TYPE "LIOLink_3UG4825_typeParam"
TITLE = LIOLink_3UG4825_typeParam
VERSION : 0.1
// Data set (index) 131 (parameters)
   STRUCT
      reserved : Array[0..15] of Byte;   // Reserved
      groupDiagnostics : Bool := TRUE;   // Group diagnostics: Default: true, false; disabled, true: enabled
      groupErrorDiagnostics : Bool := TRUE;   // Group error diagnostics: Default: true, false; disabled, true: enabled
      reserved1 : Bool;   // Reserved
      reserved2 : Bool;   // Reserved
      localLimitChange : Bool := TRUE;   // Local threshold change: Default: true, false; disabled, true: enabled
      localParameterChange : Bool := TRUE;   // Local parameter change: Default: true, false; disabled, true: enabled
      localReset : Bool := TRUE;   // Local reset: Default: true, false; disabled, true: enabled
      retentiveErrorMemory : Bool;   // Retentive error memory: Default: false, false; disabled, true: enabled
      analogValueCoding : Byte := 16#0E;   // Analog value coding: Default: 14, Min: 0(disabled), Max: 255
      reserved3 : Array[18..23] of Byte;   // Reserved
      resetResponse : Byte := 16#01;   // Reset response: Default: 16#01, 16#00: manual, 16#01: automatic
      delayOn : Bool := TRUE;   // ON-delay time (at Power ON): Default: true, false: disabled, true: enabled
      delayOn0 : Bool;   // False
      delayReset : Bool := TRUE;   // ON-delay time (at manual reset): Default: true, false: disabled, true: enabled
      delayReset0 : Bool;   // False
      delayRestart : Bool;   // ON-delay time (at restart): Default: true, false: disabled, true: enabled
      delayRestart0 : Bool;   // False
      reserved4 : Bool;   // Reserved
      reserved5 : Bool;   // Reserved
      delayTime : Int;   // ON-delay time: Resolution: 0.1=1s, Default: 0s, Min: 0.1s or 0s (disabled), Max: 999.9s
      delayTimeTripUp : Int;   // Tripping delay time (in the case of current overshoot): Resolution: 0.1s=1, Default: 0, Min: 0.1s or 0s, Max: 999.9s
      reserved6 : Word;   // Reserved
      tresholdUp : Int := 100;   // Threshold for overshoot: Resolution: 0.01A=1, Default: 1A, Min: 0.03A, Max: 40A
      reserved9 : Word;   // Reserved
      warningTresholdUp : Int := 50;   // Warning threshold for overshoot: Resolution: 0.01A=1, Default: 0,5A, Min: 0.03A or 0A (disabled), Max: 40A
      reserved7 : Array[38..43] of Byte;   // Reserved
      hysteresis : Int := 5;   // Hysteresis: Resolution: Resolution: 1%=1, Default: 5%, Min: 5% or 0% (disabled), Max: 50%
      reserved10 : Byte;   // Reserved
      responseRelay : Byte;   // Relay switching response: Default: 16#00, 16#00: Closed-circuit principle NC, 16#01: Open-circuit principle NO
   END_STRUCT;
END_TYPE

TYPE "LIOLink_3UG4825_typeAll"
TITLE = LIOLink_3UG4825_typeAll
VERSION : 0.1
// Contains all the information about 3UG4825
   STRUCT
      parameterPage0 : "LIOLink_typeParameterPage0";   // ID0: Parameter page 0
      systemCommands : Byte;   // ID2: System Commands (0x80 for device reset, 0x82 for factory reset)
      vendorName : String[11];   // ID16: Vendor name
      vendorText : String[64];   // ID17: Vendor text
      productName : String[64];   // ID18: Product name
      productID : String[14];   // ID19: Product ID
      serialNumber : String[16];   // ID21: Serial number
      hwRevision : String[7];   // ID22: Hardware revision
      fwRevision : String[7];   // ID23: Firmware revision
      appSpecificName : String[32];   // ID24: Application specific name
      diagnostics : "LIOLink_3UG4825_typeDiag";   // ID92: Diagnostics
      measuredValues : "LIOLink_3UG4825_typeMeasure";   // ID94: Measurement values
      parameters : "LIOLink_3UG4825_typeParam";   // ID131: Parameters
   END_STRUCT;
END_TYPE

TYPE "LIOLink_3UG4825_typeDiag"
TITLE = LIOLink_3UG4825_typeDiag
VERSION : 0.1
// Data set (index) 92 - diagnostics
   STRUCT
      reserved : Array[0..15] of Byte;   // Reserved
      ready : Bool;   // Ready
      groupError : Bool;   // Group error
      groupWarning : Bool;   // Group warning
      reserved1 : Bool;   // Reserved
      reserved2 : Bool;   // Reserved
      parameterAssign : Bool;   // Parameter assignment active
      parameterInvalid : Bool;   // Invalid parameter
      internalError : Bool;   // Self-test error/internal error
      reserved3 : Byte;   // Reserved
      errorNumber : Word;   // Parameter error number
      reserved4 : Array[20..25] of Byte;   // Reserved
      delayTimeRunning : Bool;   // ON-delay time running
      delayLevelUp : Bool;   // Tripping delay time running (threshold for overshoot)
      reserved5 : Bool;   // Reserved
      initTimeRunning : Bool;   // Initialization time running after applying the control supply voltage
      reserved6 : Bool;   // Reserved
      reserved7 : Bool;   // Reserved
      reserved8 : Bool;   // Reserved
      reserved9 : Bool;   // Reserved
      levelUp : Bool;   // Threshold for overshoot exceeded
      reserved10 : Bool;   // Reserved
      warningLevelUp : Bool;   // Warning threshold for overshoot exceeded
      reserved11 : Bool;   // Reserved
      reserved12 : Bool;   // Reserved
      reserved13 : Bool;   // Reserved
      reserved14 : Bool;   // Reserved
      reserved15 : Bool;   // Reserved
      wireBreak : Bool;   // Wire break
      shortCircuit : Bool;   // Short-circuit
      rangeOvershoot : Bool;   // Measuring range overshoot
      reserved16 : Bool;   // Reserved
      reserved17 : Bool;   // Reserved
      reserved18 : Bool;   // Reserved
      reserved19 : Bool;   // Reserved
      reserved20 : Bool;   // Reserved
      reserved21 : Byte;   // Reserved
   END_STRUCT;
END_TYPE

// folder: LIOLink/Common/Device-specific data types/SIRIUS/SIRIUS 3UG48/3UG4832

TYPE "LIOLink_3UG4832_typeMeasure"
TITLE = LIOLink_3UG4832_typeMeasure
VERSION : 0.1
// Contains measured value dataset of 3UG4832
   STRUCT
      reserved : Array[0..15] of Byte;   // Reserved
      voltageU1 : Word;   // Voltage
      reserved1 : Array[18..27] of Byte;   // Reserved
   END_STRUCT;
END_TYPE

TYPE "LIOLink_3UG4832_typeParam"
TITLE = LIOLink_3UG4832_typeParam
VERSION : 0.1
// LIOLink_3UG4851_typeParam
   STRUCT
      reserved : Array[0..15] of Byte;   // Reserved
      groupDiagnostics : Bool := TRUE;   // Group diagnostics: Default: true, false; disabled, true: enabled
      groupErrorDiagnostics : Bool := TRUE;   // Group error diagnostics: Default: true, false; disabled, true: enabled
      reserved1 : Bool;   // Reserved
      reserved2 : Bool;   // Reserved
      localLimitChange : Bool := TRUE;   // Local threshold change: Default: true, false; disabled, true: enabled
      localParameterChange : Bool := TRUE;   // Local parameter change: Default: true, false; disabled, true: enabled
      localReset : Bool := TRUE;   // Local reset: Default: true, false; disabled, true: enabled
      retentiveErrorMemory : Bool;   // Retentive error memory: Default: false, false; disabled, true: enabled
      analogValueCoding : Byte := 16#2C;   // Analog value coding: Default: 44, Min: 0(disabled), Max: 255
      reserved3 : Array[18..23] of Byte;   // Reserved
      resetResponse : Byte := 16#01;   // Reset response: Default: 16#01, 16#00: manual, 16#01: automatic
      delayOn : Bool := TRUE;   // ON-delay time (at Power ON): Default: true, false: disabled, true: enabled
      delayOn0 : Bool;   // False
      delayReset : Bool := TRUE;   // ON-delay time (at manual reset): Default: true, false: disabled, true: enabled
      delayReset0 : Bool;   // False
      reserved6 : Bool;   // Reserved
      reserved9 : Bool;   // Reserved
      reserved4 : Bool;   // Reserved
      reserved5 : Bool;   // Reserved
      delayTime : Int := 0;   // ON-delay time: Resolution: 0.1=1s, Default: 0s, Min: 0.1s or 0s (disabled), Max: 999.9s
      delayTimeTripUp : Int;   // Tripping delay time (in the case of voltage overshoot): Resolution: 0.1s=1, Default: 0, Min: 0.1s or 0s, Max: 999.9s
      delayTimeTripDown : Int;   // Tripping delay time (in the case of voltage undershoot): Resolution: 0.1s=1, Default: 0, Min: 0.1s or 0s, Max: 999.9s
      tresholdUp : Int := 3000;   // Threshold for overshoot: Resolution: 0.1V=1, Default: 300, Min: 10V or 0V (disabled), Max: 600V
      tresholdDown : Int := 2000;   // Threshold for undershoot: Resolution: 0.1V=1, Default: 200, Min: 10V or 0V (disabled), Max: 600V
      warningTresholdUp : Int := 3000;   // Warning threshold for overshoot: Resolution: 0.1V=1, Default: 300, Min: 10V or 0V (disabled), Max: 600V
      warningTresholdDown : Int := 2000;   // Warning threshold for undershoot: Resolution: 0.1V=1, Default: 200, Min: 10V or 0V (disabled), Max: 600V
      reserved7 : Array[40..43] of Byte;   // Reserved
      hysteresis : Int := 50;   // Hysteresis: Resolution: 0.1V=1, Default: 5V, Min: 0.1V or 0V (disabled), Max: 300V
      responseRelay : Byte;   // Relay switching response: Default: 16#00, 16#00: Closed-circuit principle NC, 16#01: Open-circuit principle NO
      reserved8 : Byte;   // Reserved
   END_STRUCT;
END_TYPE

TYPE "LIOLink_3UG4832_typeDiag"
TITLE = LIOLink_3UG4832_typeDiag
VERSION : 0.1
// Data set (index) 92 - diagnostics
   STRUCT
      reserved : Array[0..15] of Byte;   // Reserved
      ready : Bool;   // Read
      groupError : Bool;   // Group error
      groupWarning : Bool;   // Group warning
      reserved1 : Bool;   // Reserved
      reserved2 : Bool;   // Reserved
      parameterAssign : Bool;   // Parameter assignment active
      parameterInvalid : Bool;   // Invalid parameter
      internalError : Bool;   // Self-test error/internal error
      reserved3 : Byte;   // Reserved
      errorNumber : Word;   // Parameter error number
      reserved4 : Array[20..25] of Byte;   // Reserved
      delayTimeRunning : Bool;   // ON-delay time running
      delayLevelUp : Bool;   // Tripping delay time running (threshold for overshoot)
      delayLevelDown : Bool;   // Tripping delay time running (threshold for undershoot)
      reserved5 : Bool;   // Reserved
      reserved6 : Bool;   // Reserved
      reserved7 : Bool;   // Reserved
      reserved8 : Bool;   // Reserved
      reserved9 : Bool;   // Reserved
      levelUp : Bool;   // Threshold for overshoot exceeded
      levelDown : Bool;   // Threshold for undershoot violated
      warningLevelUp : Bool;   // Warning threshold for overshoot exceeded
      warningLevelDown : Bool;   // Warning threshold for undershoot violated
      reserved10 : Bool;   // Reserved
      reserved11 : Bool;   // Reserved
      reserved12 : Bool;   // Reserved
      reserved13 : Bool;   // Reserved
   END_STRUCT;
END_TYPE

TYPE "LIOLink_3UG4832_typeAll"
TITLE = LIOLink_3UG4832_typeAll
VERSION : 0.1
// Contains all the information about 3UG4832
   STRUCT
      parameterPage0 : "LIOLink_typeParameterPage0";   // ID0: Parameter page 0
      systemCommands : Byte;   // ID2: System Commands (0x80 for device reset, 0x82 for factory reset)
      vendorName : String[11];   // ID16: Vendor name
      vendorText : String[64];   // ID17: Vendor text
      productName : String[64];   // ID18: Product name
      productID : String[14];   // ID19: Product ID
      hwRevision : String[7];   // ID22: Hardware revision
      fwRevision : String[7];   // ID23: Firmware revision
      appSpecificName : String[32];   // ID24: Application specific name
      diagnostics : "LIOLink_3UG4832_typeDiag";   // ID92: Diagnostics
      measuredValues : "LIOLink_3UG4832_typeMeasure";   // ID94: Measurement values
      parameters : "LIOLink_3UG4832_typeParam";   // ID131: Parameters
   END_STRUCT;
END_TYPE

// folder: LIOLink/Common/Device-specific data types/SIRIUS/SIRIUS 3UG48/3UG4841

TYPE "LIOLink_3UG4841_typeMeasure"
TITLE = LIOLink_3UG4841_typeMeasure
VERSION : 0.1
// Data set (index) 94 (measured values)
   STRUCT
      reserved : Array[0..15] of Byte;   // Reserved
      valueCosPhiPa : Word;   // Cos Phi Value (PA) Min:0 Max:0,99
      currentActivePa : Word;   // Active current Ir/Ires (PA) Min:0,2A Max:10A
      currentApparentPa : Word;   // Apparent current Is (PA) Min:0,2A Max:10A
      voltageActivePa : Word;   // Active voltage U (PA) Min:30V Max:690V
      powerActivePa : Word;   // Active power Pw (PA) Min:6W Max:6900W
      reserved1 : Array[26..29] of Byte;   // Reserved
      currentActive : DWord;   // Active current Ir/Ires (PA) Min:0,2A Max:10A
      currentApparent : DWord;   // Apparent current Is Min:0,2A Max:10A
      powerActive : DWord;   // Active power Pw Min:6W Max:6900W
      reserved2 : Array[42..49] of Byte;   // Reserved
   END_STRUCT;
END_TYPE

TYPE "LIOLink_3UG4841_typeParam"
TITLE = LIOLink_3UG4841_typeParam
VERSION : 0.1
// Data set (index) 131 (parameters)
   STRUCT
      reserved : Array[0..15] of Byte;   // Reserved
      groupDiagnostics : Bool := TRUE;   // Group diagnostics: Default: true, false; disabled, true: enabled
      groupErrorDiagnostics : Bool := TRUE;   // Group error diagnostics: Default: true, false; disabled, true: enabled
      reserved1 : Bool;   // Reserved
      reserved2 : Bool;   // Reserved
      localLimitChange : Bool := TRUE;   // Local threshold change: Default: true, false; disabled, true: enabled
      localParameterChange : Bool := TRUE;   // Local parameter change: Default: true, false; disabled, true: enabled
      localReset : Bool := TRUE;   // Local reset: Default: true, false; disabled, true: enabled
      retentiveErrorMemory : Bool;   // Retentive error memory: Default: false, false; disabled, true: enabled
      analogValueCoding : Byte := 16#2B;   // Analog value coding: Default: 43, Min: 0(disabled), Max: 255
      reserved3 : Array[18..23] of Byte;   // Reserved
      resetResponse : Byte := 16#01;   // Reset response: Default: 16#01, 16#00: manual, 16#01: automatic
      delayOn : Bool := TRUE;   // ON-delay time (at Power ON): Default: true, false: disabled, true: enabled
      delayOn0 : Bool;   // False
      delayReset : Bool := TRUE;   // ON-delay time (at manual reset): Default: true, false: disabled, true: enabled
      delayReset0 : Bool;   // False
      delayRestart : Bool;   // ON-delay time (at restart): Default: true, false: disabled, true: enabled
      delayRestart0 : Bool;   // False
      reserved4 : Bool;   // Reserved
      reserved5 : Bool;   // Reserved
      delayTime : Int;   // ON-delay time: Resolution: 0.1=1s, Default: 0s, Min: 0.1s or 0s (disabled), Max: 999.9s
      delayTimeCosPhiTripUp : Int;   // Tripping delay time (in the case of overshoot of the cos phi value): Resolution: 0.1s=1, Default: 0, Min: 0.1s or 0s, Max: 999.9s
      delayTimeCosPhiTripDown : Int;   // Tripping delay time (in the case of undershoot of the cos phi value): Resolution: 0.1s=1, Default: 0, Min: 0.1s or 0s, Max: 999.9s
      delayTimeCurrentTripUp : Int;   // Tripping delay time (in the case of active current overshoot): Resolution: 0.1s=1, Default: 0, Min: 0.1s or 0s, Max: 999.9s
      delayTimeCurrentTripDown : Int;   // Tripping delay time (in the case of active current undershoot): Resolution: 0.1s=1, Default: 0, Min: 0.1s or 0s, Max: 999.9s
      tresholdCosPhiUp : Byte := 16#32;   // Threshold for overshoot of the cos phi value: Resolution: 0.01=1, Default: 0.5, Min: 0.01 or 0 (disabled), Max: 0.99
      tresholdCosPhiDown : Byte := 16#14;   // Threshold for undershoot of the cos phi value: Resolution: 0.01=1, Default: 0.2, Min: 0.01 or 0 (disabled), Max: 0.99
      tresholdCurrentUp : DInt := 30;   // Threshold for overshoot of the active current value: Resolution: 0.1A=1, Default: 3A, Min: 0.2A or 0A (disabled), Max: 10A
      tresholdCurrentDown : DInt := 10;   // Threshold for undershoot of the active current value: Resolution: 0.1A=1, Default: 1A, Min: 0.2A or 0A (disabled), Max: 10A
      warningTresholdCosPhiUp : Byte := 16#32;   // Warning threshold for overshoot: Resolution: 0.01A=1, Default: 2.5A, Min: 0.05A or 0A (disabled), Max: 10A
      warningTresholdCosPhiDown : Byte := 16#14;   // Warning threshold for undershoot: Resolution: 0.01A=1, Default: 1.5A, Min: 0.05A or 0A (disabled), Max: 10A
      warningTresholdCurrentUp : DInt := 30;   // Warning threshold for overshoot of the active current value: Resolution: 0.1A=1, Default: 3A, Min: 0.2A or 0A (disabled), Max: 10A
      warningTresholdCurrentDown : DInt := 10;   // Warning threshold for undershoot of the active current value: Resolution: 0.1A=1, Default: 1A, Min: 0.2A or 0A (disabled), Max: 10A
      reserved6 : Array[56..65] of Byte;   // Reserved
      hysteresisCosPhi : Byte := 16#0A;   // Hysteresis (cos phi): Resolution: 0.01=1, Default: 0.1, Min: 0.1 or 0 (disabled), Max: 0.2
      reserved7 : Byte;   // Reserved
      hysteresisCurrent : DInt := 5;   // Hysteresis (active current): Resolution: 0.1A=1, Default: 0,5A, Min: 0.1A or 0A (disabled), Max: 3A
      responseRelay : Byte;   // Relay switching response: Default: 16#00, 16#00: Closed-circuit principle NC, 16#01: Open-circuit principle NO
      reserved8 : Byte;   // Reserved
   END_STRUCT;
END_TYPE

TYPE "LIOLink_3UG4841_typeDiag"
TITLE = LIOLink_3UG4841_typeDiag
VERSION : 0.1
// Data set (index) 92 - diagnostics
   STRUCT
      reserved : Array[0..15] of Byte;   // Reserved
      ready : Bool;   // Ready
      groupError : Bool;   // Group error
      groupWarning : Bool;   // Group warning
      reserved1 : Bool;   // Reserved
      reserved2 : Bool;   // Reserved
      parameterAssign : Bool;   // Parameter assignment active
      parameterInvalid : Bool;   // Invalid parameter
      internalError : Bool;   // Self-test error/internal error
      reserved3 : Byte;   // Reserved
      errorNumber : Word;   // Parameter error number
      reserved4 : Array[20..25] of Byte;   // Reserved
      delayTimeRunning : Bool;   // ON-delay time running
      delayCosPhiUp : Bool;   // Tripping delay time running (threshold for overshoot: cos phi value)
      delayLCosPhiDown : Bool;   // Tripping delay time running (threshold for undershoot: cos phi value)
      delayCurrentUp : Bool;   // Tripping delay time running (threshold for overshoot: active current value)
      delayCurrentDown : Bool;   // Tripping delay time running (threshold for undershoot: active current value)
      reserved5 : Bool;   // Reserved
      reserved6 : Bool;   // Reserved
      reserved7 : Bool;   // Reserved
      cosPhiUp : Bool;   // Threshold value for overshoot exceeded (cos phi value)
      cosPhiDown : Bool;   // Threshold value for undershoot violated (cos phi value)
      currentUp : Bool;   // Threshold for overshoot exceeded (active current value)
      currentDown : Bool;   // Threshold for undershoot violated (active current value)
      warningCosPhiUp : Bool;   // Warning threshold for overshoot exceeded (cos phi value)
      warningCosPhiDown : Bool;   // Warning threshold for undershoot violated (cos phi value)
      warningCurrentUp : Bool;   // Warning threshold for overshoot exceeded (active current value)
      warningCurrentDown : Bool;   // Warning threshold for undershoot violated (active current value)
      reserved8 : Word;   // Reserved
   END_STRUCT;
END_TYPE

TYPE "LIOLink_3UG4841_typeAll"
TITLE = LIOLink_3UG4841_typeAll
VERSION : 0.1
// Contains all the information about 3UG4841
   STRUCT
      parameterPage0 : "LIOLink_typeParameterPage0";   // ID0: Parameter page 0
      systemCommands : Byte;   // ID2: System Commands (0x80 for device reset, 0x82 for factory reset)
      vendorName : String[11];   // ID16: Vendor name
      vendorText : String[64];   // ID17: Vendor text
      productName : String[64];   // ID18: Product name
      productID : String[14];   // ID19: Product ID
      hwRevision : String[7];   // ID22: Hardware revision
      fwRevision : String[7];   // ID23: Firmware revision
      appSpecificName : String[32];   // ID24: Application specific name
      diagnostics : "LIOLink_3UG4841_typeDiag";   // ID92: Diagnostics
      measuredValues : "LIOLink_3UG4841_typeMeasure";   // ID94: Measurement values
      parameters : "LIOLink_3UG4841_typeParam";   // ID131: Parameters
   END_STRUCT;
END_TYPE

// folder: LIOLink/Common/Device-specific data types/SIRIUS/SIRIUS 3UG48/3UG4851

TYPE "LIOLink_3UG4851_typeMeasure"
TITLE = LIOLink_3UG4851_typeMeasure
VERSION : 0.1
// Data set (index) 94 (measured values)
   STRUCT
      reserved : Array[0..15] of Byte;   // Reserved
      speed : Word;   // Speed Min:0 Max:2200
   END_STRUCT;
END_TYPE

TYPE "LIOLink_3UG4851_typeDiag"
TITLE = LIOLink_3UG4851_typeDiag
VERSION : 0.1
// Data set (index) 92 - diagnostics
   STRUCT
      reserved : Array[0..15] of Byte;   // Reserved
      ready : Bool;   // Ready
      groupError : Bool;   // Group error
      groupWarning : Bool;   // Group warning
      reserved1 : Bool;   // Reserved
      reserved2 : Bool;   // Reserved
      parameterAssign : Bool;   // Parameter assignment active
      parameterInvalid : Bool;   // Invalid parameter
      internalError : Bool;   // Self-test error/internal error
      reserved3 : Byte;   // Reserved
      errorNumber : Word;   // Parameter error number
      reserved4 : Array[20..25] of Byte;   // Reserved
      delayTimeRunning : Bool;   // ON-delay time running
      delayLevelUp : Bool;   // Tripping delay time running (threshold for overshoot)
      delayLevelDown : Bool;   // Tripping delay time running (threshold for undershoot)
      reserved5 : Bool;   // Reserved
      reserved6 : Bool;   // Reserved
      reserved7 : Bool;   // Reserved
      reserved8 : Bool;   // Reserved
      reserved9 : Bool;   // Reserved
      levelUp : Bool;   // Threshold for overshoot exceeded
      levelDown : Bool;   // Threshold for undershoot violated
      warningLevelUp : Bool;   // Warning threshold for overshoot exceeded
      warningLevelDown : Bool;   // Warning threshold for undershoot violated
      reserved10 : Bool;   // Reserved
      reserved11 : Bool;   // Reserved
      reserved12 : Bool;   // Reserved
      reserved13 : Bool;   // Reserved
      rangeOvershoot : Bool;   // Sensor - Measuring range overshoot
      reserved14 : Bool;   // Reserved
      reserved15 : Bool;   // Reserved
      reserved16 : Bool;   // Reserved
      reserved17 : Bool;   // Reserved
      reserved18 : Bool;   // Reserved
      reserved19 : Bool;   // Reserved
      reserved20 : Bool;   // Reserved
      reserved21 : Byte;   // Reserved
   END_STRUCT;
END_TYPE

TYPE "LIOLink_3UG4851_typeParam"
TITLE = LIOLink_3UG4851_typeParam
VERSION : 0.1
// Data set (index) 131 (parameters)
   STRUCT
      reserved : Array[0..15] of Byte;   // Reserved
      groupDiagnostics : Bool := TRUE;   // Group diagnostics: Default: true, false; disabled, true: enabled
      groupErrorDiagnostics : Bool := TRUE;   // Group error diagnostics: Default: true, false; disabled, true: enabled
      reserved1 : Bool;   // Reserved
      reserved2 : Bool;   // Reserved
      localLimitChange : Bool := TRUE;   // Local threshold change: Default: true, false; disabled, true: enabled
      localParameterChange : Bool := TRUE;   // Local parameter change: Default: true, false; disabled, true: enabled
      localReset : Bool := TRUE;   // Local reset: Default: true, false; disabled, true: enabled
      retentiveErrorMemory : Bool;   // Retentive error memory: Default: false, false; disabled, true: enabled
      analogValueCoding : Byte := 16#0D;   // Analog value coding: Default: 13, Min: 0(disabled), Max: 255
      reserved3 : Array[18..23] of Byte;   // Reserved
      resetResponse : Byte := 16#01;   // Reset response: Default: 16#01, 16#00: manual, 16#01: automatic
      delayOn : Bool := TRUE;   // ON-delay time (at Power ON): Default: true, false: disabled, true: enabled
      delayOn0 : Bool;   // False
      delayReset : Bool := TRUE;   // ON-delay time (at manual reset): Default: true, false: disabled, true: enabled
      delayReset0 : Bool;   // False
      reserved4 : Bool;   // Reserved
      reserved5 : Bool;   // Reserved
      reserved6 : Bool;   // Reserved
      reserved7 : Bool;   // Reserved
      delayTime : Int;   // ON-delay time: Resolution: 0.1=1s, Default: 0s, Min: 0.1s or 0s (disabled), Max: 999.9s
      delayTimeTripUp : Int;   // Tripping delay time (in the case of speed overshoot): Resolution: 0.1s=1, Default: 0, Min: 0.1s or 0s, Max: 999.9s
      delayTimeTripDown : Int;   // Tripping delay time (in the case of speed undershoot): Resolution: 0.1s=1, Default: 0, Min: 0.1s or 0s, Max: 999.9s
      tresholdUp : Int := 1400;   // Threshold for speed overshoot: Default: 1400rpm, Min: 0.1rpm or 0rpm (disabled), Max: 2200rpm
      tresholdDown : Int := 800;   // Threshold for speed undershoot: Default: 800rpm, Min: 0.1rpm or 0rpm (disabled), Max: 2200rpm
      warningTresholdUp : Int := 1400;   // Warning threshold for speed overshoot: Default: 1400rpm, Min: 0.1rpm or 0rpm (disabled), Max: 2200rpm
      warningTresholdDown : Int := 800;   // Warning threshold for speed undershoot: Default: 800rpm, Min: 0.1rpm or 0rpm (disabled), Max: 2200rpm
      reserved8 : Array[40..43] of Byte;   // Reserved
      hysteresis : Int := 50;   // Hysteresis: Resolution: 0.1=1, Default: 5, Min: 0.1 or 0 (disabled), Max: 99.9
      responseRelay : Byte;   // Relay switching response: Default: 16#00, 16#00: Closed-circuit principle NC, 16#01: Open-circuit principle NO
      reserved9 : Byte;   // Reserved
   END_STRUCT;
END_TYPE

TYPE "LIOLink_3UG4851_typeAll"
TITLE = LIOLink_3UG4851_typeAll
VERSION : 0.1
// Contains all the information about 3UG4851
   STRUCT
      parameterPage0 : "LIOLink_typeParameterPage0";   // ID0: Parameter page 0
      systemCommands : Byte;   // ID2: System Commands (0x80 for device reset, 0x82 for factory reset)
      vendorName : String[11];   // ID16: Vendor name
      vendorText : String[64];   // ID17: Vendor text
      productName : String[64];   // ID18: Product name
      productID : String[14];   // ID19: Product ID
      hwRevision : String[7];   // ID22: Hardware revision
      fwRevision : String[7];   // ID23: Firmware revision
      appSpecificName : String[32];   // ID24: Application specific name
      diagnostics : "LIOLink_3UG4851_typeDiag";   // ID92: Diagnostics
      measuredValues : "LIOLink_3UG4851_typeMeasure";   // ID94: Measurement values
      parameters : "LIOLink_3UG4851_typeParam";   // ID131: Parameters
   END_STRUCT;
END_TYPE

// folder: LIOLink/Common/Device-specific data types/SIRIUS/SIRIUS WD

TYPE "LIOLink_8WD46_typeAll"
TITLE = LIOLink_8WD46_typeAll
// Contains all the information about 8WD46
   STRUCT
      systemCommand : Byte;   // system command to reset to default settings
      vendorName : String[48];   // Siemens AG (default)
      vendorText : String[48];   // http://www.siemens.com/io-link (default)
      productName : String[32];   // 8WD46 IO-Link 9 Segments (default)
      productId : String[16];   // 8WD4613-5HH47 (default)
      productText : String[64];   // SIRIUS Signaling Column 8WD46 IO-Link (default)
      serialNumber : String[16];   // 0000000000000000 (default)
      hwRevision : String[16];   // 1.0 (default)
      fwRevision : String[16];   // 1.2.0 (default)
      appSpecificName : String[32];   // *** (default)
      functionTag : String[32];   // *** (default)
      locationTag : String[32];   // *** (default)
      deviceStatus : Byte;   // device status
      deviceStatusDetailed : Byte;   // detailed device status
      opHour : DWord;   // operation time in hours
      operatingMode : Byte;   // operating mode (signal mode, auto scale mode, ...)
      lightEffects : Array[1..15] of "LIOLink_8WD46_typeLightEffects";   // optical effects of each segment (1 to 9/15)
      soundMode : Array[1..10] of "LIOLink_8WD46_typeSoundMode";   // sound effects (10 configurable)
      powerReduction : Byte;   // power reduction (0: on / 1: off)
      fillLevelMode : Byte;   // only in level mode (0: use settings of segment 1-9,15 / 1: use settings of segment 1 )
      headlong : Byte;   // orientation of installation (normal / overhead)
      elementCount : Byte;   // number of elements
   END_STRUCT;
END_TYPE

TYPE "LIOLink_8WD46_typeLightEffects"
TITLE = LIOLink_8WD46_typeLightEffects
// Light Effect data record
   STRUCT
      effect : Byte;   // light effect (permanet light, flash, ...)
      pwmR : Byte;   // Red component (only relevant for individual color PWM)
      pwmG : Byte;   // Green component (only relevant for individual color PWM)
      pwmB : Byte;   // Blue component (only relevant for individual color PWM)
      brightness : Byte;   // brightness of the segmenttt
      defaultColor : Byte;   // default color (0: individual color PWM, 1: red, 2: green, ...)
      reserved : Byte;   // reserved
      priority : Byte;   // priority in auto scale mode
   END_STRUCT;
END_TYPE

TYPE "LIOLink_8WD46_typeSoundMode"
TITLE = LIOLink_8WD46_typeSoundMode
// Sound Mode data record
   STRUCT
      mode : Byte;   // tone type (0: off, 1: Continuous tone, 2: pulse tone, ...)
      frequency1Start : Word;   // Frequency at the start of a cycle in Hz
      frequency2Stop : Word;   // Frequency at the end of a cycle in Hz
      frequency1Periode : Word;   // Frequency for time betwen frequency 1 and 2 in Hz*10
      volume : Byte;   // 0: low, 1: mediummm, 2: loud, 3: very loud
      count : Word;   // repeat count
      brakeToRepeat : Word;   // Pause after repeat
      BrakeBetweenCycles : Word;   // Duration of the pause beween cycle in ms
      holdingPeriodeFrequency2 : Word;   // Setting of thehold time for full-scale frequency in ms
   END_STRUCT;
END_TYPE

// folder: LIOLink/Devices/SIRIUS/3RS2x

TYPE "LIOLink_3RS2_typePIQ"
TITLE = 3RS14_PIQ
VERSION : 0.1
   STRUCT
      startOnDlyTime : Bool;   // Start ON-delay time / Starte Anlaufverzögerungszeit
      res0 : Bool;   // reserved / Reserviert
      res1 : Bool;   // reserved / Reserviert
      reset : Bool;   // Reset
      res2 : Bool;   // reserved / Reserviert
      res3 : Bool;   // reserved / Reserviert
      res4 : Bool;   // reserved / Reserviert
      res5 : Bool;   // reserved / Reserviert
      res6 : Bool;   // reserved / Reserviert
      res7 : Bool;   // reserved / Reserviert
      res8 : Bool;   // reserved / Reserviert
      res9 : Bool;   // reserved / Reserviert
      res10 : Bool;   // reserved / Reserviert
      res11 : Bool;   // reserved / Reserviert
      res12 : Bool;   // reserved / Reserviert
      res13 : Bool;   // reserved / Reserviert
   END_STRUCT;
END_TYPE

TYPE "LIOLink_3RS2_typePII"
TITLE = 3RS14_PII
VERSION : 0.1
   STRUCT
      ready : Bool;   // Ready / Betriebsbereit
      res0 : Bool;   // reserved / Reserviert
      groupError : Bool;   // Group error / Sammelfehler
      groupWarning : Bool;   // General or group warning / Sammelwarnung
      statusK1 : Bool;   // Status output relay K1; 1: 14NO/11C closed and 12NC/11C open, 0: 12NC/11C closed and 14NO/11C open / Status Ausgangrelais K1
      statusK2 : Bool;   // Status output relay K2; 1: 24NO/21C closed and 22NC/21C open, 0: 22NC/21C closed and 24NO/21C open / Status Ausgangrelais K2
      statusK3 : Bool;   // Status output relay K3; 1: 33NO/34NO closed, 0: 33NO/34NO open / Status Ausgangrelais K3
      res1 : Bool;   // reserved / Reserviert
      analogValueCoding : Byte;   // Analog value coding bits 0 to 4 / Analogwertcodierung (nur Bit 0..4)
      AnalogValue : Int;   // Analog value / Analogwert
   END_STRUCT;
END_TYPE

// folder: LIOLink/Devices/SIRIUS/3SU1/3SU1 Electronic Module

TYPE "LIOLink_3SU1_ElecModule_typePII"
VERSION : 0.1
   STRUCT
      reserved : DWord;
      status : Byte;
      input0 : Bool;
      input1 : Bool;
      input2 : Bool;
      input3 : Bool;
      input4 : Bool;
      input5 : Bool;
      input6 : Bool;
      input7 : Bool;
   END_STRUCT;
END_TYPE

TYPE "LIOLink_3SU1_ElecModule_typePIQ"
VERSION : 0.1
   STRUCT
      res0 : DWord;   // Reserved
      output0 : Bool;
      output1 : Bool;
      output2 : Bool;
      output3 : Bool;
      output4 : Bool;
      output5 : Bool;
      output6 : Bool;
      output7 : Bool;
      res1 : Byte;   // Reserved
   END_STRUCT;
END_TYPE

// folder: LIOLink/Profiles

TYPE "LIOLink_typeIdentificationObjects"
   STRUCT
      vendorID : Word;   // Vendor ID
      deviceID : DWord;   // Device ID
      vendorName : String[64];   // Vendor name
      vendorText : String[64];   // Vendor text
      productName : String[64];   // Product name
      productID : String[64];   // Product ID
      productText : String[64];   // Product text
      serialNumber : String[16];   // Serial number
      hwRevision : String[64];   // Hardware revision
      fwRevision : String[64];   // Firmware revision
      appSpecificTag : String[32];   // Application specific name
      locationTag : String[32];   // Location tag
      functionTag : String[32];   // Function tag
   END_STRUCT;
END_TYPE

// folder: Base blocks

FUNCTION_BLOCK "LIOLink_Master"   // FB5002, SCL
TITLE = LIOLink_Master
{ S7_Optimized_Access := 'FALSE' }
AUTHOR : SIOS
FAMILY : LIOLink
VERSION : 4.0
// Backs up or restores the complete configuration of Siemens IO-Link master modules
   VAR_INPUT
      execute : Bool;   // Request to execute function
      logicalAddr : DInt;   // Logical address of IO-Link master module (sub module for ET 200eco PN)
      mode : Int;   // 0: backup, 1: restore
   END_VAR
   VAR_OUTPUT
      done : Bool;   // TRUE: Commanded functionality has been completed successfully
      busy : Bool;   // TRUE: FB is not finished and new output values can be expected
      error : Bool;   // TRUE: An error occurred during the execution of the FB
      status : Word := 16#7000;   // 16#0000 - 16#7FFF: Status of the FB, 16#8000 - 16#FFFF: Error identification
      diagnostics : "LIOLink_typeDiagnostics";   // Diagnostics information of FB
      len : DInt;   // Total length of parameter record (number of bytes)
   END_VAR
   VAR_IN_OUT
      record : Array[0..#UPPER_LIMIT_8_PORT] of Byte;   // Record to store backup in or restore from
   END_VAR
   VAR
      statExecuteOld : Bool;   // Old value of 'execute' input for edge detection
      statDone : Bool;   // Static value for output 'done'
      statBusy : Bool;   // Static value for output 'busy'
      statError : Bool;   // Static value for output 'error'
      statStatus : Word := 16#7000;   // Static value for output 'status'
      statStatusBits AT statStatus : Array[0..15] of Bool;
      statSubfunctionStatus : DWord;   // Status or return value of called FBs, FCs and system blocks
      statFBErrorState : Int;   // State in the state machine of the block where the error occurred
      statFBState : Int := 0;   // State in the state machine of the FB
      statEmptyDiagnostics : "LIOLink_typeDiagnostics";   // Empty diagnostics information (for initialization purposes only)
      instRdRec : RDREC;   // System function "read data record"
      instWrRec : WRREC;   // System function "write data record"
      statRecStruct : Struct   // structured database for different jobs of RDREC/WRREC
         reset : Struct   // structure of data record for reset (NEW)
            ExtendedFunctionNum : Byte;   // extended function number (01=PUSH, 02=PULL)
            Options : Byte;   // options, not used
            SequenceNo : DWord;   // sequence number (please see manual)
            payload : Array[0..233] of Byte;   // payload data (raw data)
         END_STRUCT;
         backup : Struct   // structure of data record for backup (NEW)
            ExtendedFunctionNum : Byte;   // extended function number (01=PUSH, 02=PULL)
            Options : Byte;   // options, not used
            SequenceNo : DWord;   // sequence number (please see manual)
            payload : Array[0..233] of Byte;   // payload data (raw data)
         END_STRUCT;
         restore : Struct   // structure of data record for restore (NEW)
            ExtendedFunctionNum : Byte;   // extended function number (01=PUSH, 02=PULL)
            Options : Byte;   // options, not used
            SequenceNo : DWord;   // sequence number (please see manual)
            payload : Array[0..233] of Byte;   // payload data (raw data)
         END_STRUCT;
      END_STRUCT;
      statLogicalAddr : DWord;   // Static value for input 'logicalAddress'
      statMode : Int;   // Static value for input 'mode'
      statSegment : DInt;   // current segment
      statAddress : DInt;   // current address
      statLen : DInt;   // total length of operated data
   END_VAR
   VAR_TEMP
      tempExecute : Bool;   // Temporary value for input 'execute'
      tempIndex : DInt;   // loop index
      tempLen : Int;   // current length of data record
   END_VAR
   VAR CONSTANT
      UPPER_LIMIT_4_PORT : DInt := 10239;   // Upper limit of data record array for 4 port master
      UPPER_LIMIT_8_PORT : DInt := 17549;   // Upper limit of data record array for 8 port master
      INDEX : Int := 120;   // Index of data record for backup/restore operations
      MODE_BACKUP : Int := 0;   // Mode backup
      MODE_RESTORE : Int := 1;   // Mode restore
      FUNC_PUSH : Byte := 16#01;   // Extended function number for push
      FUNC_PULL : Byte := 16#02;   // Extended function number for pull
      LEN_HEADER : Int := 6;   // Length of header
      MAX_SIZE_SEGMENT : Int := 234;   // Max. 234 Byte per segment
      FB_STATE_NO_PROCESSING : Int := 0;   // FB state: No processing
      FB_STATE_RESET : Int := 1;   // FB state: reset (essential before each backup/restore operation)
      FB_STATE_BACKUP : Int := 11;   // FB state: backup
      FB_STATE_RESTORE : Int := 21;   // FB state: restore segment data
      FB_STATE_VERIFY : Int := 22;   // FB state: verify restore
      STATUS_EXECUTION_FINISHED : Word := 16#0000;   // Execution finished without errors
      STATUS_NO_CALL : Word := 16#7000;   // No job being currently processed
      STATUS_FIRST_CALL : Word := 16#7001;   // First call after incoming new job (rising edge 'execute')
      STATUS_SUBSEQUENT_CALL : Word := 16#7002;   // Subsequent call during active processing without further details
      STATUS_OFFSET_BACKUP : Word := 16#7100;   // Offset for status during backup operation
      STATUS_OFFSET_RESTORE : Word := 16#7200;   // Offset for status during restore operation
      SUB_STATUS_NO_ERROR : Word := 16#0000;   // No error occured in subfunction call
      ERR_UNKNOWN_MODULE : Word := 16#80B0;   // unknown type of module, check subfunctionStatus
      ERR_ARRAY_UNSUPPORTED : Word := 16#8201;   // Record array doesn't fit expected limits
      ERR_UNKNOWN_MODE : Word := 16#8202;   // Unknown mode
      ERR_SEQ_NUMBER : Word := 16#8401;   // Error: IO-Link master returned a sequence number indicating an error, see "diagnostics"
      ERR_UNDEFINED_STATE : Word := 16#8600;   // Error: due to an undefined state in state machine
      ERR_WRRC_RESET : Word := 16#8601;   // Error: WRREC encountered an error during reset, see "diagnostics"
      ERR_RDREC_BACKUP : Word := 16#8602;   // Error: RDREC encountered an error during backup, see "diagnostics"
      ERR_WRREC_RESTORE : Word := 16#8603;   // Error: WRREC encountered an error during restore, see "diagnostics"
      ERR_RDREC_VERIFY : Word := 16#8604;   // Error: RDREC encountered an error during verification of restore, see "diagnostics"
      ERR_UNKNOWN_RECORD : DWord := 16#DF80_B000;   // Error: Data record not known in module
      SEQ_NUM_RESET : DWord := 16#FFFF_FFFF;   // Sequence number for reset before backup/restore operations
      SEQ_NUM_RESTORE_ONGOING : DWord := 16#FFFF_FF01;   // Sequence number: restore ongoing
      SEQ_NUM_ACTIVATION_ONGOING : DWord := 16#FFFF_FF02;   // Sequence number: activation ongoing
      SEQ_NUM_ACTIVATION_DONE : DWord := 16#FFFF_FF03;   // Sequence number: activation done
      SEQ_NUM_CRC_FAILED : DWord := 16#FFFF_FF04;   // Sequence number: CRC check failed
      SEQ_NUM_BLOB_INVALID : DWord := 16#FFFF_FF05;   // Sequence number: blob data invalid
      SEQ_NUM_WRONG_SEQUENCE : DWord := 16#FFFF_FF06;   // Sequence number: wrong sequence number
      SEQ_NUM_WRONG_SIZE : DWord := 16#FFFF_FF07;   // Sequence number: wrong data record size
   END_VAR
BEGIN
   REGION BLOCK INFO HEADER
     //===============================================================================
     // Siemens / (c)Copyright 2020
     //-------------------------------------------------------------------------------
     // Title:            LIOLink_Master
     // Function:         Backs up or restores the complete configuration of Siemens IO-Link master modules
     // Library:          LIOLink
     // Author:           Siemens Industry Online Support
     // Tested with:      CPU 315-2 PN/DP FW 3.2
     // Engineering:      TIA Portal V16
     // Restrictions:     --
     // Requirements:     One of the following IO-Link master modules:
     //                   - ET 200SP, CM 4x IO-Link 6ES7137-6BD00-0BA0 FW V2.2.0 or higher
     //                   - ET 200AL, CM 4x IO-Link 6ES7147-5JD00-0BA0 FW V1.1.0 or higher
     //                   - ET 200pro, EM 4 IO-Link 6ES7147-4JD00-0AB0 FW V1.0.0 or higher
     //                   - ET 200eco PN, IO-Link Master 6ES7148-6JD00-0AB0 FW V1.0.0 or higher
     //                   - ET 200eco PN, CM 8x IO-Link 6ES7148-6JG00-0BB0 FW V1.0.0 or higher
     //                   - S7-1500, CM 8xIO-Link 6ES7547-1JF00-0AB0 FW V1.0.0 or higher
     //-------------------------------------------------------------------------------
     // Change log table:
     // Version  | Date       | Expert in charge       | Changes applied
     //----------|------------|------------------------|------------------------------
     // 01.00.00 | 28.02.2015 | SUP Applications       | First release
     // 02.00.00 | 30.09.2016 | SUP Applications       | Integration of complete backup/restore for master and device parameter (new ET 200eco PN)
     // 03.00.00 | 30.09.2017 | SUP Applications       | Reduction to use only one way for complete backup/restore of master and device parameter
     // 03.00.01 | 14.12.2018 | SUP Applications       | Renamed function block from IO_LINK_MASTER to IO_LINK_MASTER_4. No functional changes
     // 04.00.00 | 01.09.2020 | Online Support         | Implemented Programming styleguide for S7-1200/1500 and PLCopen
     //                                                | Combined FBs for 4 Port and 8 Port IO-Link Masters to one FB
     //                                                | Renamed FB to LIOLink_Master
     //===============================================================================
   END_REGION

   #tempExecute := #execute; // Work with temporary value / create process image

   REGION TRIGGERING
     IF (#tempExecute = TRUE) AND (#statExecuteOld = FALSE)
       AND (#statStatus = #STATUS_NO_CALL)
     THEN // First call; initialize FB
       #statDone := FALSE;
       #statBusy := TRUE;
       #statError := FALSE;
       #statStatus := #STATUS_FIRST_CALL;
       #statSubfunctionStatus := #SUB_STATUS_NO_ERROR;
       #statFBErrorState := 0;
       #diagnostics := #statEmptyDiagnostics;

       // Save input parameters
       #statLogicalAddr := DINT_TO_DWORD(#logicalAddr);
       #statMode := #mode;

       // Initialize internal tags 
       #statSegment := 0;
       #statAddress := 0;
       #statLen := 0;

       IF #statMode = #MODE_BACKUP THEN
         FOR #tempIndex := 0 TO #UPPER_LIMIT_8_PORT DO   // initialize data record before backup
           #record[#tempIndex] := 16#0;
         END_FOR;
         #statFBState := #FB_STATE_RESET;
       ELSIF #statMode = #MODE_RESTORE THEN
         #statFBState := #FB_STATE_RESET;
       ELSE
         #statStatus := #ERR_UNKNOWN_MODE;
       END_IF;

     ELSIF (#statStatus = #STATUS_FIRST_CALL) THEN
       #statStatus := #STATUS_SUBSEQUENT_CALL;
     END_IF;

     // Edge detection 'execute' input
     #statExecuteOld := #tempExecute;
   END_REGION TRIGGERING

   REGION STATE_MACHINE
     CASE #statFBState OF
       #FB_STATE_NO_PROCESSING:
         REGION no processing
           ; // No processing active
         END_REGION no processing

       #FB_STATE_RESET:
         REGION reset
           #statRecStruct.reset.ExtendedFunctionNum := #FUNC_PUSH;
           #statRecStruct.reset.SequenceNo := #SEQ_NUM_RESET;  // reset save/restore operations

           #instWrRec(REQ    := true,
                      ID     := #statLogicalAddr,
                      INDEX  := #INDEX,
                      LEN    := #LEN_HEADER,
                      RECORD := #statRecStruct.reset);

           IF #instWrRec.DONE = TRUE THEN
             #instWrRec(REQ := FALSE); // Reset request

             IF #statMode = #MODE_BACKUP THEN
               #statFBState := #FB_STATE_BACKUP;
             ELSE
               #statFBState := #FB_STATE_RESTORE;
             END_IF;
           ELSIF #instWrRec.ERROR = TRUE AND #instWrRec.STATUS = #ERR_UNKNOWN_RECORD THEN
             #statStatus := #ERR_UNKNOWN_MODULE; // set status = unknown type of module
             #statSubfunctionStatus := #instWrRec.STATUS;
             #statFBErrorState := #statFBState;
           ELSIF #instWrRec.ERROR = TRUE THEN
             #statStatus := #ERR_WRRC_RESET;
             #statSubfunctionStatus := #instWrRec.STATUS;
             #statFBErrorState := #statFBState;
           END_IF;
         END_REGION reset

       #FB_STATE_BACKUP:
         REGION backup
           #instRdRec(REQ    := TRUE,
                      ID     := #statLogicalAddr,
                      INDEX  := #INDEX,
                      MLEN   := #LEN_HEADER + #MAX_SIZE_SEGMENT,
                      RECORD := #statRecStruct.backup);

           // evaluation of RDREC
           IF #instRdRec.VALID = TRUE THEN
             IF #instRdRec.LEN > #LEN_HEADER AND #statRecStruct.backup.ExtendedFunctionNum = #FUNC_PULL THEN
               #statStatus := #STATUS_OFFSET_BACKUP OR DWORD_TO_BYTE(#statRecStruct.backup.SequenceNo);  // append segment number
               #statSegment := DWORD_TO_DINT(#statRecStruct.backup.SequenceNo);
               #tempLen := #instRdRec.LEN - #LEN_HEADER;

               // store payload
               FOR #tempIndex := 0 TO #tempLen - 1 DO
                 #record[#statAddress + #tempIndex] := #statRecStruct.backup.payload[#tempIndex];
               END_FOR;

               // add total length of data
               #statLen := #statLen + #tempLen;

               // set pointer to next entry in parameter blob
               #statAddress := #statAddress + #tempLen;

             ELSIF #instRdRec.LEN = #LEN_HEADER THEN
               // Reset request
               #instRdRec(REQ    := FALSE,
                          RECORD := #statRecStruct.backup);

               #statStatus := #STATUS_EXECUTION_FINISHED;
             END_IF;

           ELSIF #instRdRec.ERROR = TRUE THEN
             #statStatus := #ERR_RDREC_BACKUP;
             #statSubfunctionStatus := #instRdRec.STATUS;
             #statFBErrorState := #statFBState;
             #statLen := #instRdRec.LEN;
           END_IF;
         END_REGION backup

       #FB_STATE_RESTORE:
         REGION restore
           // load restore data segment from parameter blob (max. 234 Byte per segment)
           IF #instWrRec.BUSY = FALSE AND #instWrRec.DONE = FALSE THEN // Writing hasn't started
             #statRecStruct.restore.ExtendedFunctionNum := #FUNC_PUSH;
             #statRecStruct.restore.SequenceNo := DINT_TO_DWORD(#statSegment); // sequence number
             #statStatus := #STATUS_OFFSET_RESTORE OR DWORD_TO_BYTE(#statRecStruct.restore.SequenceNo);

             // load segment data = payload
             FOR #tempIndex := 0 TO #MAX_SIZE_SEGMENT - 1 DO
               #statRecStruct.restore.payload[#tempIndex] := #record[#statAddress + #tempIndex];
             END_FOR;
           END_IF;

           // write segment data
           #instWrRec(REQ    := TRUE,
                      ID     := #statLogicalAddr,
                      INDEX  := #INDEX,
                      LEN    := #LEN_HEADER + #MAX_SIZE_SEGMENT,
                      RECORD := #statRecStruct.restore);

           IF #instWrRec.DONE = TRUE THEN
             #statLen := #statLen + #MAX_SIZE_SEGMENT;
             #instWrRec(REQ := FALSE); // Reset request
             #statFBState := #FB_STATE_VERIFY;
           ELSIF #instWrRec.ERROR = TRUE THEN
             #statStatus := #ERR_WRREC_RESTORE;
             #statSubfunctionStatus := #instWrRec.STATUS;
             #statFBErrorState := #statFBState;
           END_IF;
         END_REGION restore

       #FB_STATE_VERIFY: // Verify restore
         REGION verify
           #instRdRec(REQ    := TRUE,
                      ID     := #statLogicalAddr,
                      INDEX  := #INDEX,
                      MLEN   := #LEN_HEADER + #MAX_SIZE_SEGMENT,
                      RECORD := #statRecStruct.backup);

           IF #instRdRec.VALID = TRUE AND #statRecStruct.backup.ExtendedFunctionNum = #FUNC_PULL THEN
             IF #statRecStruct.backup.SequenceNo = #SEQ_NUM_RESTORE_ONGOING
               OR #statRecStruct.backup.SequenceNo = #SEQ_NUM_ACTIVATION_ONGOING
             THEN
               #statSegment := #statSegment + 1;
               #statAddress := #statAddress + #MAX_SIZE_SEGMENT;

               // Reset request
               #instRdRec(REQ    := FALSE,
                          RECORD := #statRecStruct.backup);

               #statFBState := #FB_STATE_RESTORE;
             ELSIF #statRecStruct.backup.SequenceNo = #SEQ_NUM_ACTIVATION_DONE THEN //
               // Reset request
               #instRdRec(REQ    := FALSE,
                          RECORD := #statRecStruct.backup);

               #statStatus := #STATUS_EXECUTION_FINISHED;
             ELSIF #statRecStruct.backup.SequenceNo = #SEQ_NUM_CRC_FAILED
               OR #statRecStruct.backup.SequenceNo = #SEQ_NUM_BLOB_INVALID
               OR #statRecStruct.backup.SequenceNo = #SEQ_NUM_WRONG_SEQUENCE
               OR #statRecStruct.backup.SequenceNo = #SEQ_NUM_WRONG_SIZE
             THEN
               #statStatus := #ERR_SEQ_NUMBER;
               #statSubfunctionStatus := #statRecStruct.backup.SequenceNo;
               #statFBErrorState := #statFBState;
             END_IF;
           ELSIF #instRdRec.ERROR = TRUE THEN
             #statStatus := #ERR_RDREC_VERIFY;
             #statSubfunctionStatus := #instRdRec.STATUS;
             #statFBErrorState := #statFBState;
           END_IF;
         END_REGION verify

       ELSE // Undefined state in state machine reached
         REGION undefined state
           #statStatus := #ERR_UNDEFINED_STATE;
         END_REGION undefined state no relevant case, ready for new request
     END_CASE;
   END_REGION

   REGION OUTPUTS
     // Write outputs
     IF (#statStatus = #STATUS_EXECUTION_FINISHED) AND (#statDone = FALSE) THEN // Execution finished without errors
       REGION execution finished
         #statDone := TRUE;
         #statBusy := FALSE;
         #statError := FALSE;
         #len := #statLen;
         // execution aborted --> set state no processing
         #statFBState := #FB_STATE_NO_PROCESSING;
       END_REGION execution finished

     ELSIF (#statStatusBits[7] = TRUE) AND (#statError = FALSE) THEN // Error occurred (#statStatus is 16#8000 to 16#FFFF)
       REGION error occured
         #statDone := FALSE;
         #statBusy := FALSE;
         #statError := TRUE;
         // Write diagnostics
         #diagnostics.status := #statStatus;
         #diagnostics.subfunctionStatus := #statSubfunctionStatus;
         #diagnostics.stateNumber := #statFBErrorState;
         // Call instructions with FALSE to be ready for next job
         #instRdRec(REQ    := FALSE,
                    RECORD := #statRecStruct.backup);

         #instWrRec(REQ := FALSE);
         // execution aborted --> set state no processing
         #statFBState := #FB_STATE_NO_PROCESSING;
       END_REGION error occured

     ELSIF (#tempExecute = FALSE) AND ((#statDone = TRUE) OR (#statError = TRUE)) THEN // Reset outputs
       REGION execute reset
         #statDone := FALSE;
         #statBusy := FALSE;
         #statError := FALSE;
         #statStatus := #STATUS_NO_CALL;
         #len := 0;
       END_REGION execute reset
     END_IF;

     REGION write static values to outputs
       #done := #statDone;
       #busy := #statBusy;
       #error := #statError;
       #status := #statStatus;
       ENO := NOT #statError;
     END_REGION write static values to outputs
   END_REGION OUTPUTS
END_FUNCTION_BLOCK

FUNCTION_BLOCK "LIOLink_Device"   // FB5003, SCL
TITLE = LIOLink_Device
{ S7_Optimized_Access := 'FALSE' }
AUTHOR : SIOS
FAMILY : LIOLink
VERSION : 4.0
// Acyclically reads or writes data records from and to IO-Link devices
   VAR_INPUT
      execute : Bool;   // Request to execute function / Request Function / Neuer Auftrag
      logicalAddr : DInt;   // Logical address of IO-Link master module (sub module for ET 200eco PN) / Hardwarekennung des IOL-Master Moduls (HW_IO) aus HW-Konfiguration
      cap : Int := 227;   // Client Access Point; 0xB400 for ET 200eco PN, CM 8x IO-Link, else 0xE003 (227) / Client Access Point (CAP), bei ET200 immer 227 dez
      readWrite : Bool;   // FALSE: read, TRUE: write / Lese und Schreibzugriff auf IO-Link Device 0: Lesen, 1: schreiben
      port : Int;   // Port on IO-Link master module / Port/ Kanalnummer an dem das IO-Link Device betrieben wird. (ET200 = 0 .. 4)
      index : Int;   // Address parameter index (IO-Link device); 0..32767: IOL-D; 65535: port functions / Adressparameter Index (IO-Link Device) 0..32767 IOL-D, 65535 port functions
      subindex : Int;   // Address parameter subindex (IO-Link device); 0: full record; 1-255: single parameter / Adressparameter Subindex (IO-Link Device) 0 ges. Record; 1-255 einz. Parameter
      writeLen : Int;   // Length of writing data (net data) / Länge der zu schreibenden Daten (Nettodaten)
      timeout : Time := T#20s;   // Time after which the request is aborted
   END_VAR
   VAR_OUTPUT
      done : Bool;   // TRUE: Commanded functionality has been completed successfully / Gültigkeit 0: Daten nicht gültig; 1: Daten gültig
      busy : Bool;   // TRUE: FB is not finished and new output values can be expected / 0: Auftrag abgeschlossen 1: Auftrag in Bearbeitung
      error : Bool;   // TRUE: An error occurred during the execution of the FB / Fehler Flag 0: kein Fehler; 1: Abbruch der Funktion mit Fehler
      status : Word := 16#7000;   // 16#0000-16#7FFF: Status of the FB, 16#8000-16#FFFF: Error identification / IO-Link Fehlerstatus; ERROR Flag = 1 - detaillierte IO-Link Fehlerstatus
      diagnostics : "LIOLink_typeDiagnostics";   // Diagnostics information of FB
      readLen : Int;   // Length of read data record (number of bytes) / Länge des gelesenen Datensatzes (Anzahl Bytes)
   END_VAR
   VAR_IN_OUT
      record : Array[0..#UPPER_LIMIT] of Byte;   // Data area for reading/writing data (max. 232 byte) / Datenbereich für LESEN / SCHREIBEN (max. 232 Byte)
   END_VAR
   VAR
      statExecuteOld : Bool;   // Old value of 'execute' input for edge detection
      statDone : Bool;   // Static value for output 'done'
      statBusy : Bool;   // Static value for output 'busy'
      statError : Bool;   // Static value for output 'error'
      statStatus : Word := 16#7000;   // Static value for output 'status'
      statStatusBits AT statStatus : Array[0..15] of Bool;
      statSubfunctionStatus : DWord;   // Status of WRREC/RDREC or error code from IO-Link Master (%W1: IO-Link Master error, %W0: ISDU error)
      statSubfunctionStatusBytes AT statSubfunctionStatus : Array[0..3] of Byte;
      statFBErrorState : DInt;   // State in the state machine of the block where the error occurred
      statFBState : DInt := 0;   // State in the state machine of the FB
      statEmptyDiagnostics : "LIOLink_typeDiagnostics";   // Empty diagnostics information (for initialization purposes only)
      instRdRec : RDREC;   // System function "read data record" / Funktion Datensatz lesen (ehemals SFB52)
      instWrRec : WRREC;   // System function "write data record" / Funktion Datensatz schreiben (ehemals SFB53)
      instPoll : TP;   // poll rate read data record / Pollzeit für "Datensatz lesen"
      instMonitor : TON;   // request monitoring time / Überwachungszeit für Aufträge
      statRead : Struct   // data area for reading data / Datenbereich für Lesedaten
         header : Struct   // Header
            call : Struct   // Header for read/write data record / header for read/write data record
               extFunctionNum : Byte := 16#8;   // Extended function number (fix coded 0x08) / extended function number (fix coded 08h)
               port : Byte;   // variable port (user interface) 0...255
               fiIndex : Word := 16#FE4A;   // FI index (fix coded 65098)
            END_STRUCT;
            IOL : Struct   // Header for IO-Link / header for IO-Link
               control : Byte;   // Control byte; 0x03: read, 0x02: write / RD_WR = 0 = read = Control:=0x03 / / RD_WR = 1 = write = Control:=0x02
               indexHighByte : Byte;   // index of data record 0…32767 (high byte)
               indexLowByte : Byte;   // index of data record 0…32767 (low byte)
               subindex : Byte;   // subindex for data record 0...255
            END_STRUCT;
         END_STRUCT;
         data : Array[0..231] of Byte;   // User data
      END_STRUCT;
      statWrite : Struct   // data area for writing data / Datenbereich für Schreibdaten
         header : Struct   // Header
            call : Struct   // Header for read/write data record / header for read/write data record
               extFunctionNum : Byte := 16#8;   // Extended function number (fix coded 0x08) / extended function number (fix coded 08h)
               port : Byte;   // Variable port (user interface) 0...255 / variable port (user interface) 0...255
               fiIndex : Word := 16#FE4A;   // FI index (fix coded 65098)
            END_STRUCT;
            IOL : Struct   // Header for IO-Link / header for IO-Link
               control : Byte;   // Control byte; 0x03: read, 0x02: write / RD_WR = 0 = read = Control:=0x03 / / RD_WR = 1 = write = Control:=0x02
               indexHighByte : Byte;   // index of data record 0…32767 (high byte)
               indexLowByte : Byte;   // index of data record 0…32767 (low byte)
               subindex : Byte;   // subindex for data record 0...255
            END_STRUCT;
         END_STRUCT;
         data : Array[0..231] of Byte;   // User data
      END_STRUCT;
      statLogicalAddr : DWord;   // Static value for input 'logicalAddr'
      statCap : Int;   // Static value for input 'cap'
      statReadWrite : Bool;   // Stativ value for input 'readWrite'
      statTimeout : Time;   // Static value for input 'timeout'
      statLen : Int;   // Length of data to be written to device
   END_VAR
   VAR_TEMP
      tempExecute : Bool;   // Temporary value for input 'execute'
      tempIndex : DInt;   // run tag for counting loops / Laufvariable für for-Schleifen
   END_VAR
   VAR CONSTANT
      MODE_READ : Bool := FALSE;   // Mode to read data
      MODE_WRITE : Bool := TRUE;   // Mode to write data
      MAX_PORT : Int := 63;   // Max. possible port
      MAX_INDEX : Int := 32767;   // Max. possible index
      INDEX_PORT_FUNC : DInt := 65535;   // Index to address port functions
      MAX_SUBINDEX : Int := 255;   // Max. possible subindex
      MAX_DATA : Int := 232;   // Max. size of data to be transferred
      UPPER_LIMIT : Int := 231;   // Upper limit of data to be transferred
      POLLING_PERIOD : Time := T#100ms;   // Time in between polls
      FB_STATE_NO_PROCESSING : DInt := 0;   // FB state: No processing
      FB_STATE_WRITE : Int := 1;   // Write data record
      FB_STATE_POLL : Int := 2;   // wait and poll for response
      LEN_HEADER : Int := 8;   // Length of header
      CONTROL_WRITE : Byte := 16#02;   // Write data record
      CONTROL_READ : Byte := 16#03;   // Read data record
      STATUS_EXECUTION_FINISHED : Word := 16#0000;   // Execution finished without errors
      STATUS_NO_CALL : Word := 16#7000;   // No job being currently processed
      STATUS_FIRST_CALL : Word := 16#7001;   // First call after incoming new job (rising edge 'execute')
      STATUS_SUBSEQUENT_CALL : Word := 16#7002;   // Subsequent call during active processing without further details
      SUB_STATUS_NO_ERROR : Word := 16#0000;   // No error occured in subfunction call
      ERR_WRONG_PORT : Word := 16#8201;   // Error: wrong port
      ERR_WRONG_INDEX : Word := 16#8202;   // Error: wrong index
      ERR_WRONG_SUBINDEX : Word := 16#8203;   // Error: wrong subindex
      ERR_WRONG_LENGTH : Word := 16#8205;   // Error: wrong length for write data record
      ERR_IO_LINK : Word := 16#8401;   // Error: IO-Link master returned error code, see "diagnostics"
      ERR_REQUEST_TIMEOUT : Word := 16#8403;   // Error: Request timed out
      ERR_INCONSISTENT_DATA : Word := 16#8402;   // Error: Read data record doesn't match request
      ERR_UNDEFINED_STATE : Word := 16#8600;   // Error: due to an undefined state in state machine
      ERR_WRREC : Word := 16#8601;   // Error: WRREC encountered an error, see "diagnostics"
      ERR_RDREC : Word := 16#8602;   // Error: RDREC encountered an error, see "diagnostics"
      STATUS_MASK : DWord := 16#00FF_FF00;   // Mask to filter error codes
      STATUS_RESOURCE_BUSY : DWord := 16#0080_C200;   // Status from WRREC/RDREC: Resource is busy
   END_VAR
   // // diagnostics.subfunctionStatus : Status of WRREC/RDREC or error code from IO-Link Master (%W1: IO-Link Master error, %W0: ISDU error)
BEGIN
   REGION BLOCK INFO HEADER
     //===============================================================================
     // Siemens / (c)Copyright 2020
     //-------------------------------------------------------------------------------
     // Title:            LIOLink_Device
     // Function:         Acyclically reads or writes data records from and to IO-Link devices
     // Library:          LIOLink
     // Author:           Siemens Industry Online Support
     // Tested with:      CPU 315-2 PN/DP FW 3.2
     // Engineering:      TIA Portal V16
     // Restrictions:     S7-300/400
     // Requirements:     --
     //-------------------------------------------------------------------------------
     // Change log table:
     // Version  | Date       | Expert in charge       | Changes applied
     //----------|------------|------------------------|------------------------------
     // 02.00.00 | 30.09.2013 | Online Support         | First release for TIA Portal V12 SP1 as IO_LINK_CALL
     // 02.01.00 | 14.03.2014 | Online Support         | Upgrade to TIA Portal V13
     //                                                | Upgrade of system function 'WRREC' from V1.0 to V1.1
     // 03.00.00 | 28.02.2015 | SUP Applications       | Upgrade to TIA Portal V13 SP1
     //                                                | Renamed FB to IO_LINK_DEVICE 
     // 03.01.00 | 15.09.2015 | SUP Applications       | Change of #IOL_INDEX AND #Port lower boundry to 0 and improved behaviour when called in cyclic OBs with > 100 ms
     // 04.00.00 | 01.09.2020 | Online Support         | Implemented Programming styleguide for S7-1200/1500 and PLCopen
     //                                                | Renamed FB to LIOLink_Device 
     //===============================================================================
   END_REGION

   #tempExecute := #execute; // Work with temporary value / create process image

   REGION TRIGGERING
     IF (#tempExecute = TRUE) AND (#statExecuteOld = FALSE) // Check if FB is triggered
       AND (#statStatus = #STATUS_NO_CALL)
     THEN // First call; initialize FB
       #statDone := FALSE;
       #statBusy := TRUE;
       #statError := FALSE;
       #statStatus := #STATUS_FIRST_CALL;
       #statSubfunctionStatus := #SUB_STATUS_NO_ERROR;
       #statFBErrorState := 0;
       #diagnostics := #statEmptyDiagnostics;
       #readLen := 0;

       // Save input parameters
       #statLogicalAddr := DINT_TO_DWORD(#logicalAddr);
       #statCap := #cap;
       #statReadWrite := #readWrite;
       #statTimeout := #timeout;

       // Initialize data area
       #statRead.header."call"."port" := 16#0;
       #statRead.header.IOL.indexLowByte := 16#0;
       #statRead.header.IOL.indexHighByte := 16#0;
       #statRead.header.IOL.subindex := 16#0;
       #tempIndex := 0; // initialize loop counter      
       FOR #tempIndex := 0 TO #UPPER_LIMIT DO
         #statWrite.data[#tempIndex] := 16#0;
         #statRead.data[#tempIndex] := 16#0;
       END_FOR;

       // Check parameters
       IF (#port < 0) OR (#port > #MAX_PORT) THEN
         #statStatus := #ERR_WRONG_PORT;
       ELSIF (#index < 0) OR (#index > #MAX_INDEX AND #index <> #INDEX_PORT_FUNC) THEN
         #statStatus := #ERR_WRONG_INDEX;
       ELSIF (#subindex < 0) OR (#subindex > #MAX_SUBINDEX) THEN
         #statStatus := #ERR_WRONG_SUBINDEX;
       ELSIF #statReadWrite = #MODE_WRITE AND (#writeLen < 1 OR #writeLen > #MAX_DATA) THEN
         #statStatus := #ERR_WRONG_LENGTH;
       END_IF;

       // setup call header
       #statWrite.header."call"."port" := INT_TO_BYTE(#port);

       // setup IOL header 
       #statWrite.header.IOL.indexLowByte := INT_TO_BYTE(#index);
       #statWrite.header.IOL.indexHighByte := WORD_TO_BYTE(SHR(IN := INT_TO_WORD(#index), N := 8));
       #statWrite.header.IOL.subindex := INT_TO_BYTE(#subindex);

       // BODY (data max. 232 Byte, Array 0..231 of Byte) 
       IF #statReadWrite = #MODE_WRITE THEN // Write data record requested, copy data from "record"
         #statWrite.header.IOL.control := #CONTROL_WRITE;
         #statLen := #writeLen + #LEN_HEADER; // data length header + data = IO-Link write data record
         // copy "record" to working area
         FOR #tempIndex := 0 TO #writeLen - 1 DO
           #statWrite.data[#tempIndex] := #record[#tempIndex];
         END_FOR;
       ELSE // Read data record requested
         // Empty record array
         FOR #tempIndex := 0 TO #UPPER_LIMIT DO
           #record[#tempIndex] := 16#0;
         END_FOR;

         #statWrite.header.IOL.control := #CONTROL_READ;
         #statLen := #LEN_HEADER; // data length only header = IO-Link read data record
       END_IF;

       IF #statStatus = #STATUS_FIRST_CALL THEN // Parameters OK
         #statFBState := #FB_STATE_WRITE;  // Start sequence
       END_IF;

     ELSIF (#statStatus = #STATUS_FIRST_CALL) THEN
       #statStatus := #STATUS_SUBSEQUENT_CALL;
     END_IF;

     // Edge detection 'execute' input
     #statExecuteOld := #tempExecute;
   END_REGION TRIGGERING

   REGION STATE_MACHINE
     CASE #statFBState OF
       #FB_STATE_NO_PROCESSING:
         REGION no processing
           ; // No processing active
         END_REGION no processing

       #FB_STATE_WRITE:
         REGION write
           // To read data records, the IO-Link master modules needs to know which port is required. Therefore it is necessary
           // to send at first a request via write data record (header, 8 byte). As response the IO-Link master module will 
           // send the required data record.

           #instWrRec(REQ    := TRUE,
                      ID     := #statLogicalAddr,
                      INDEX  := #statCap,
                      LEN    := #statLen,
                      RECORD := #statWrite);

           IF #instWrRec.ERROR THEN
             IF (#instWrRec.STATUS AND #STATUS_MASK) = #STATUS_RESOURCE_BUSY THEN
               #instWrRec(REQ := FALSE); // Reset requeset
             ELSE
               #statStatus := #ERR_WRREC;
               #statSubfunctionStatus := #instWrRec.STATUS;
               #statFBErrorState := #statFBState;
             END_IF;
           ELSIF #instWrRec.DONE = TRUE THEN
             #instWrRec(REQ := FALSE); // Reset requeset

             #statFBState := #FB_STATE_POLL;
           END_IF;
         END_REGION write

       #FB_STATE_POLL: // wait and poll for response
         REGION poll
           #instPoll(IN := TRUE,
                     PT := #POLLING_PERIOD);

           // read data record on falling edge
           #instRdRec(REQ    := NOT #instPoll.Q,
                      ID     := #statLogicalAddr,
                      INDEX  := #statCap,
                      MLEN   := #MAX_DATA,
                      RECORD := #statRead);

           IF #instRdRec.ERROR = TRUE THEN
             IF (#instRdRec.STATUS AND #STATUS_MASK) = #STATUS_RESOURCE_BUSY THEN
               // Reset requests and try again
               #instPoll(IN := FALSE,
                         PT := #POLLING_PERIOD);

               #instRdRec(REQ    := FALSE,
                          RECORD := #statRead);
             ELSE
               #statStatus := #ERR_RDREC;
               #statSubfunctionStatus := #instRdRec.STATUS;
               #statFBErrorState := #statFBState;
             END_IF;
           ELSIF #instRdRec.VALID THEN
             IF // check the response wether it matches the request (compare PORT, INDEX and SUBINDEX)
               (#statWrite.header."call"."port" <> #statRead.header."call"."port")
               OR (#statWrite.header.IOL.indexHighByte <> #statRead.header.IOL.indexHighByte)
               OR (#statWrite.header.IOL.indexLowByte <> #statRead.header.IOL.indexLowByte)
               OR (#statWrite.header.IOL.subindex <> #statRead.header.IOL.subindex)
             THEN // read data record doesn't match the request
               #statStatus := #ERR_INCONSISTENT_DATA;  // output status no consistent data
             ELSIF #statRead.header.IOL.control = B#16#80 THEN // check the response for IO-Link errors
               // State 0x80 = IOL_CALL_RES PDU shows IO-Link error detect
               #statStatus := #ERR_IO_LINK;
               #statSubfunctionStatusBytes[0] := #statRead.data[0]; // IO-Link master error code
               #statSubfunctionStatusBytes[1] := #statRead.data[1]; // IO-Link master error code
               #statSubfunctionStatusBytes[2] := #statRead.data[2]; // ISDU error code
               #statSubfunctionStatusBytes[3] := #statRead.data[3]; // ISDU additional code
               #statFBErrorState := #statFBState;
             ELSE // read data is valid
               IF #statReadWrite = #MODE_READ THEN
                 #readLen := #instRdRec.LEN - #LEN_HEADER;
                 // only data will be output
                 FOR #tempIndex := 0 TO #instRdRec.LEN - #LEN_HEADER - 1 DO
                   #record[#tempIndex] := #statRead.data[#tempIndex];
                 END_FOR;
               END_IF;

               // Reset requests
               #instRdRec(REQ    := FALSE,
                          RECORD := #statRead);

               #instPoll(IN := FALSE,
                         PT := #POLLING_PERIOD);

               #statStatus := #STATUS_EXECUTION_FINISHED;  // request finished
             END_IF;
           END_IF;
         END_REGION poll

       ELSE // Undefined state in state machine reached
         REGION undefined state
           #statStatus := #ERR_UNDEFINED_STATE;
         END_REGION undefined state no relevant case, ready for new request
     END_CASE;
   END_REGION

   REGION MONITORING
     #instMonitor(IN := #statBusy,
                  PT := #statTimeout);

     IF #instMonitor.Q THEN
       #statStatus := #ERR_REQUEST_TIMEOUT; // request time out
     END_IF;
   END_REGION

   REGION OUTPUTS
     // Write outputs
     IF (#statStatus = #STATUS_EXECUTION_FINISHED) AND (#statDone = FALSE) THEN // Execution finished without errors
       REGION execution finished
         #statDone := TRUE;
         #statBusy := FALSE;
         #statError := FALSE;
         // execution aborted --> set state no processing
         #statFBState := #FB_STATE_NO_PROCESSING;
       END_REGION execution finished

     ELSIF (#statStatusBits[7] = TRUE) AND (#statError = FALSE) THEN // Error occurred (#statStatus is 16#8000 to 16#FFFF)
       REGION error occured
         #statDone := FALSE;
         #statBusy := FALSE;
         #statError := TRUE;
         // Write diagnostics
         #diagnostics.status := #statStatus;
         #diagnostics.subfunctionStatus := #statSubfunctionStatus;
         #diagnostics.stateNumber := #statFBErrorState;
         // Call instructions with FALSE to be ready for next job
         #instWrRec(REQ := FALSE);

         #instRdRec(REQ    := FALSE,
                    RECORD := #statRead);

         #instPoll(IN := FALSE,
                   PT := #POLLING_PERIOD);

         // execution aborted --> set state no processing
         #statFBState := #FB_STATE_NO_PROCESSING;
       END_REGION error occured

     ELSIF (#tempExecute = FALSE) AND ((#statDone = TRUE) OR (#statError = TRUE)) THEN // Reset outputs
       REGION execute reset
         #statDone := FALSE;
         #statBusy := FALSE;
         #statError := FALSE;
         #statStatus := #STATUS_NO_CALL;
         #readLen := 0;
       END_REGION execute reset
     END_IF;

     REGION write static values to outputs
       #done := #statDone;
       #busy := #statBusy;
       #error := #statError;
       #status := #statStatus;
       ENO := NOT #statError;
     END_REGION write static values to outputs
   END_REGION OUTPUTS
END_FUNCTION_BLOCK

FUNCTION_BLOCK "LIOLink_Master"   // FB50005, SCL
TITLE = LIOLink_Master / IO_LINK_MASTER
{ S7_Optimized_Access := 'TRUE' }
AUTHOR : SIOS
FAMILY : LIOLink
VERSION : 4.0
// Backs up or restores the complete configuration of Siemens IO-Link master modules / Lesen und Schreiben der Parameter für IO-Link Master Module
   VAR_INPUT
      execute : Bool;   // Request to execute function
      hwID : HW_IO;   // Hardware identifier of IO-Link master module (sub module for ET 200eco PN)
      mode : USInt;   // 0: backup, 1: restore
   END_VAR
   VAR_OUTPUT
      done : Bool;   // TRUE: Commanded functionality has been completed successfully
      busy : Bool;   // TRUE: FB is not finished and new output values can be expected
      error : Bool;   // TRUE: An error occurred during the execution of the FB
      status : Word;   // 16#0000 - 16#7FFF: Status of the FB, 16#8000 - 16#FFFF: Error identification
      diagnostics : "LIOLink_typeDiagnostics";   // Diagnostics information of FB
      len : DInt;   // Total length of parameter record (number of bytes)
   END_VAR
   VAR_IN_OUT
      record : Array[*] of Byte;   // Record to store backup in or restore from; limits for 4 Port masters: 0..10239, limits for 8 Port masters: 0..17549
   END_VAR
   VAR
      statExecuteOld : Bool;   // Old value of 'execute' input for edge detection
      statDone : Bool;   // Static value for output 'done'
      statBusy : Bool;   // Static value for output 'busy'
      statError : Bool;   // Static value for output 'error'
      statStatus : Word := 16#7000;   // Static value for output 'status'
      statSubfunctionStatus : DWord;   // Status or return value of called FBs, FCs and system blocks
      statFBErrorState : Int;   // State in the state machine of the block where the error occurred
      statFBState : Int := 0;   // State in the state machine of the FB
      statEmptyDiagnostics : "LIOLink_typeDiagnostics";   // Empty diagnostics information (for initialization purposes only)
      instRdRec : RDREC;   // System function "read data record"
      instWrRec : WRREC;   // System function "write data record"
      statRecStruct : Struct   // structured database for different jobs of RDREC/WRREC
         reset : Struct   // structure of data record for reset (NEW)
            ExtendedFunctionNum : Byte;   // extended function number (01=PUSH, 02=PULL)
            Options : Byte;   // options, not used
            SequenceNo : DWord;   // sequence number (please see manual)
            payload : Array[0..233] of Byte;   // payload data (raw data)
         END_STRUCT;
         backup : Struct   // structure of data record for backup (NEW)
            ExtendedFunctionNum : Byte;   // extended function number (01=PUSH, 02=PULL)
            Options : Byte;   // options, not used
            SequenceNo : DWord;   // sequence number (please see manual)
            payload : Array[0..233] of Byte;   // payload data (raw data)
         END_STRUCT;
         restore : Struct   // structure of data record for restore (NEW)
            ExtendedFunctionNum : Byte;   // extended function number (01=PUSH, 02=PULL)
            Options : Byte;   // options, not used
            SequenceNo : DWord;   // sequence number (please see manual)
            payload : Array[0..233] of Byte;   // payload data (raw data)
         END_STRUCT;
      END_STRUCT;
      statHwID : HW_IO;   // Static value for input 'hwID'
      statMode : USInt;   // Static value for input 'mode'
      statSegment : DInt;   // current segment
      statAddress : DInt;   // current address
      statLen : DInt;   // total length of operated data
   END_VAR
   VAR_TEMP
      tempExecute : Bool;   // Temporary value for input 'execute'
      tempLowerBound : DInt;   // Lower bound of record array
      tempUpperBound : DInt;   // Upper bound of record array
      tempIndex : DInt;   // loop index
      tempLen : UInt;   // current length of data record
   END_VAR
   VAR CONSTANT
      UPPER_LIMIT_4_PORT : DInt := 10239;   // Upper limit of data record array for 4 port master
      UPPER_LIMIT_8_PORT : DInt := 17549;   // Upper limit of data record array for 8 port master
      INDEX : USInt := 120;   // Index of data record for backup/restore operations
      MODE_BACKUP : USInt := 0;   // Mode backup
      MODE_RESTORE : USInt := 1;   // Mode restore
      FUNC_PUSH : Byte := 16#01;   // Extended function number for push
      FUNC_PULL : Byte := 16#02;   // Extended function number for pull
      LEN_HEADER : USInt := 6;   // Length of header
      MAX_SIZE_SEGMENT : UInt := 234;   // Max. 234 Byte per segment
      FB_STATE_NO_PROCESSING : Int := 0;   // FB state: No processing
      FB_STATE_RESET : Int := 1;   // FB state: reset (essential before each backup/restore operation)
      FB_STATE_BACKUP : Int := 11;   // FB state: backup
      FB_STATE_RESTORE : Int := 21;   // FB state: restore segment data
      FB_STATE_VERIFY : Int := 22;   // FB state: verify restore
      STATUS_EXECUTION_FINISHED : Word := 16#0000;   // Execution finished without errors
      STATUS_NO_CALL : Word := 16#7000;   // No job being currently processed
      STATUS_FIRST_CALL : Word := 16#7001;   // First call after incoming new job (rising edge 'execute')
      STATUS_SUBSEQUENT_CALL : Word := 16#7002;   // Subsequent call during active processing without further details
      STATUS_OFFSET_BACKUP : Word := 16#7100;   // Offset for status during backup operation
      STATUS_OFFSET_RESTORE : Word := 16#7200;   // Offset for status during restore operation
      SUB_STATUS_NO_ERROR : Word := 16#0000;   // No error occured in subfunction call
      ERR_UNKNOWN_MODULE : Word := 16#80B0;   // unknown type of module, check subfunctionStatus
      ERR_UNKNOWN_MODE : Word := 16#8200;   // Unknown mode
      ERR_ARRAY_UNSUPPORTED : Word := 16#8201;   // Record array doesn't fit expected limits
      ERR_SEQ_NUMBER : Word := 16#8401;   // Error: IO-Link master returned a sequence number indicating an error, see "diagnostics"
      ERR_UNDEFINED_STATE : Word := 16#8600;   // Error: due to an undefined state in state machine
      ERR_WRRC_RESET : Word := 16#8601;   // Error: WRREC encountered an error during reset, see "diagnostics"
      ERR_RDREC_BACKUP : Word := 16#8602;   // Error: RDREC encountered an error during backup, see "diagnostics"
      ERR_WRREC_RESTORE : Word := 16#8603;   // Error: WRREC encountered an error during restore, see "diagnostics"
      ERR_RDREC_VERIFY : Word := 16#8604;   // Error: RDREC encountered an error during verification of restore, see "diagnostics"
      ERR_UNKNOWN_RECORD : DWord := 16#DF80_B000;   // Error: Data record not known in module
      SEQ_NUM_RESET : DWord := 16#FFFF_FFFF;   // Sequence number for reset before backup/restore operations
      SEQ_NUM_RESTORE_ONGOING : DWord := 16#FFFF_FF01;   // Sequence number: restore ongoing
      SEQ_NUM_ACTIVATION_ONGOING : DWord := 16#FFFF_FF02;   // Sequence number: activation ongoing
      SEQ_NUM_ACTIVATION_DONE : DWord := 16#FFFF_FF03;   // Sequence number: activation done
      SEQ_NUM_CRC_FAILED : DWord := 16#FFFF_FF04;   // Sequence number: CRC check failed
      SEQ_NUM_BLOB_INVALID : DWord := 16#FFFF_FF05;   // Sequence number: blob data invalid
      SEQ_NUM_WRONG_SEQUENCE : DWord := 16#FFFF_FF06;   // Sequence number: wrong sequence number
      SEQ_NUM_WRONG_SIZE : DWord := 16#FFFF_FF07;   // Sequence number: wrong data record size
   END_VAR
BEGIN
   REGION BLOCK INFO HEADER
     //===============================================================================
     // Siemens / (c)Copyright 2020
     //-------------------------------------------------------------------------------
     // Title:            LIOLink_Master
     // Function:         Backs up or restores the complete configuration of Siemens IO-Link master modules
     // Library:          LIOLink
     // Author:           Siemens Industry Online Support
     // Tested with:      CPU 1513-1 PN FW 2.8
     // Engineering:      TIA Portal V16
     // Restrictions:     --
     // Requirements:     One of the following IO-Link master modules:
     //                   - ET 200SP, CM 4x IO-Link 6ES7137-6BD00-0BA0 FW V2.2.0 or higher
     //                   - ET 200AL, CM 4x IO-Link 6ES7147-5JD00-0BA0 FW V1.1.0 or higher
     //                   - ET 200pro, EM 4 IO-Link 6ES7147-4JD00-0AB0 FW V1.0.0 or higher
     //                   - ET 200eco PN, IO-Link Master 6ES7148-6JD00-0AB0 FW V1.0.0 or higher
     //                   - ET 200eco PN, CM 8x IO-Link 6ES7148-6JG00-0BB0 FW V1.0.0 or higher
     //                   - S7-1500, CM 8xIO-Link 6ES7547-1JF00-0AB0 FW V1.0.0 or higher
     //-------------------------------------------------------------------------------
     // Change log table:
     // Version  | Date       | Expert in charge       | Changes applied
     //----------|------------|------------------------|------------------------------
     // 01.00.00 | 28.02.2015 | SUP Applications       | First release
     // 02.00.00 | 30.09.2016 | SUP Applications       | Integration of complete backup/restore for master and device parameter (new ET 200eco PN)
     // 03.00.00 | 30.09.2017 | SUP Applications       | Reduction to use only one way for complete backup/restore of master and device parameter
     // 03.00.01 | 14.12.2018 | SUP Applications       | Renamed function block from IO_LINK_MASTER to IO_LINK_MASTER_4. No functional changes
     // 04.00.00 | 01.09.2020 | Online Support         | Implemented Programming styleguide for S7-1200/1500 and PLCopen
     //                                                | Combined FBs for 4 Port and 8 Port IO-Link Masters to one FB
     //                                                | Renamed FB to LIOLink_Master
     //===============================================================================
   END_REGION

   #tempExecute := #execute; // Work with temporary value / create process image

   REGION TRIGGERING
     IF (#tempExecute = TRUE) AND (#statExecuteOld = FALSE)
       AND (#statStatus = #STATUS_NO_CALL)
     THEN // First call; initialize FB
       #statDone := FALSE;
       #statBusy := TRUE;
       #statError := FALSE;
       #statStatus := #STATUS_FIRST_CALL;
       #statSubfunctionStatus := #SUB_STATUS_NO_ERROR;
       #statFBErrorState := 0;
       #diagnostics := #statEmptyDiagnostics;

       // Save input parameters
       #statHwID := #hwID;
       #statMode := #mode;

       // Initialize internal tags 
       #statSegment := 0;
       #statAddress := 0;
       #statLen := 0;

       // Check record array
       #tempLowerBound := LOWER_BOUND(ARR := #record, DIM := 1);
       #tempUpperBound := UPPER_BOUND(ARR := #record, DIM := 1);

       IF #tempLowerBound <> 0
         OR (#tempUpperBound <> #UPPER_LIMIT_4_PORT
         AND #tempUpperBound <> #UPPER_LIMIT_8_PORT)
       THEN
         #statStatus := #ERR_ARRAY_UNSUPPORTED;
       ELSE // Check mode
         IF #statMode = #MODE_BACKUP THEN
           FOR #tempIndex := 0 TO #tempUpperBound DO // initialize data record before backup
             #record[#tempIndex] := 16#0;
           END_FOR;
           #statFBState := #FB_STATE_RESET;
         ELSIF #statMode = #MODE_RESTORE THEN
           #statFBState := #FB_STATE_RESET;
         ELSE
           #statStatus := #ERR_UNKNOWN_MODE;
         END_IF;
       END_IF;

     ELSIF (#statStatus = #STATUS_FIRST_CALL) THEN
       #statStatus := #STATUS_SUBSEQUENT_CALL;
     END_IF;

     // Edge detection 'execute' input
     #statExecuteOld := #tempExecute;
   END_REGION TRIGGERING

   REGION STATE_MACHINE
     CASE #statFBState OF
       #FB_STATE_NO_PROCESSING:
         REGION no processing
           ; // No processing active
         END_REGION no processing

       #FB_STATE_RESET:
         REGION reset
           #statRecStruct.reset.ExtendedFunctionNum := #FUNC_PUSH;
           #statRecStruct.reset.SequenceNo := #SEQ_NUM_RESET;  // reset save/restore operations

           #instWrRec(REQ    := true,
                      ID     := #statHwID,
                      INDEX  := #INDEX,
                      LEN    := #LEN_HEADER,
                      RECORD := #statRecStruct.reset);

           IF #instWrRec.DONE = TRUE THEN
             #instWrRec(REQ := FALSE); // Reset request

             IF #statMode = #MODE_BACKUP THEN
               #statFBState := #FB_STATE_BACKUP;
             ELSE
               #statFBState := #FB_STATE_RESTORE;
             END_IF;
           ELSIF #instWrRec.ERROR = TRUE AND #instWrRec.STATUS = #ERR_UNKNOWN_RECORD THEN
             #statStatus := #ERR_UNKNOWN_MODULE; // set status = unknown type of module
             #statSubfunctionStatus := #instWrRec.STATUS;
             #statFBErrorState := #statFBState;
           ELSIF #instWrRec.ERROR = TRUE THEN
             #statStatus := #ERR_WRRC_RESET;
             #statSubfunctionStatus := #instWrRec.STATUS;
             #statFBErrorState := #statFBState;
           END_IF;
         END_REGION reset

       #FB_STATE_BACKUP:
         REGION backup
           #instRdRec(REQ    := TRUE,
                      ID     := #statHwID,
                      INDEX  := #INDEX,
                      MLEN   := #LEN_HEADER + #MAX_SIZE_SEGMENT,
                      RECORD := #statRecStruct.backup);

           // evaluation of RDREC
           IF #instRdRec.VALID = TRUE THEN
             IF #instRdRec.LEN > #LEN_HEADER AND #statRecStruct.backup.ExtendedFunctionNum = #FUNC_PULL THEN
               #statStatus := #STATUS_OFFSET_BACKUP OR #statRecStruct.backup.SequenceNo.%B0;  // append segment number
               #statSegment := DWORD_TO_DINT(#statRecStruct.backup.SequenceNo);
               #tempLen := #instRdRec.LEN - #LEN_HEADER;

               // store payload
               MOVE_BLK(IN    := #statRecStruct.backup.payload[0],
                        COUNT := #tempLen,
                        OUT   => #record[#statAddress]);

               // add total length of data
               #statLen := #statLen + #tempLen;

               // set pointer to next entry in parameter blob
               #statAddress := #statAddress + #tempLen;

             ELSIF #instRdRec.LEN = #LEN_HEADER THEN
               // Reset request
               #instRdRec(REQ    := FALSE,
                          RECORD := #statRecStruct.backup);

               #statStatus := #STATUS_EXECUTION_FINISHED;
             END_IF;

           ELSIF #instRdRec.ERROR = TRUE THEN
             #statStatus := #ERR_RDREC_BACKUP;
             #statSubfunctionStatus := #instRdRec.STATUS;
             #statFBErrorState := #statFBState;
             #statLen := #instRdRec.LEN;
           END_IF;
         END_REGION backup

       #FB_STATE_RESTORE:
         REGION restore
           // load restore data segment from parameter blob (max. 234 Byte per segment)
           IF #instWrRec.BUSY = FALSE AND #instWrRec.DONE = FALSE THEN // Writing hasn't started
             #statRecStruct.restore.ExtendedFunctionNum := #FUNC_PUSH;
             #statRecStruct.restore.SequenceNo := DINT_TO_DWORD(#statSegment); // sequence number
             #statStatus := #STATUS_OFFSET_RESTORE OR #statRecStruct.restore.SequenceNo.%B0;

             // load segment data = payload
             MOVE_BLK(IN    := #record[#statAddress],
                      COUNT := #MAX_SIZE_SEGMENT,
                      OUT   => #statRecStruct.restore.payload[0]);
           END_IF;

           // write segment data
           #instWrRec(REQ    := TRUE,
                      ID     := #statHwID,
                      INDEX  := #INDEX,
                      LEN    := #LEN_HEADER + #MAX_SIZE_SEGMENT,
                      RECORD := #statRecStruct.restore);

           IF #instWrRec.DONE = TRUE THEN
             #statLen := #statLen + #MAX_SIZE_SEGMENT;
             #instWrRec(REQ := FALSE); // Reset request
             #statFBState := #FB_STATE_VERIFY;
           ELSIF #instWrRec.ERROR = TRUE THEN
             #statStatus := #ERR_WRREC_RESTORE;
             #statSubfunctionStatus := #instWrRec.STATUS;
             #statFBErrorState := #statFBState;
           END_IF;
         END_REGION restore

       #FB_STATE_VERIFY: // Verify restore
         REGION verify
           #instRdRec(REQ    := TRUE,
                      ID     := #statHwID,
                      INDEX  := #INDEX,
                      MLEN   := #LEN_HEADER + #MAX_SIZE_SEGMENT,
                      RECORD := #statRecStruct.backup);

           IF #instRdRec.VALID = TRUE AND #statRecStruct.backup.ExtendedFunctionNum = #FUNC_PULL THEN
             IF #statRecStruct.backup.SequenceNo = #SEQ_NUM_RESTORE_ONGOING
               OR #statRecStruct.backup.SequenceNo = #SEQ_NUM_ACTIVATION_ONGOING
             THEN
               #statSegment := #statSegment + 1;
               #statAddress := #statAddress + #MAX_SIZE_SEGMENT;

               // Reset request
               #instRdRec(REQ    := FALSE,
                          RECORD := #statRecStruct.backup);

               #statFBState := #FB_STATE_RESTORE;
             ELSIF #statRecStruct.backup.SequenceNo = #SEQ_NUM_ACTIVATION_DONE THEN //
               // Reset request
               #instRdRec(REQ    := FALSE,
                          RECORD := #statRecStruct.backup);

               #statStatus := #STATUS_EXECUTION_FINISHED;
             ELSIF #statRecStruct.backup.SequenceNo = #SEQ_NUM_CRC_FAILED
               OR #statRecStruct.backup.SequenceNo = #SEQ_NUM_BLOB_INVALID
               OR #statRecStruct.backup.SequenceNo = #SEQ_NUM_WRONG_SEQUENCE
               OR #statRecStruct.backup.SequenceNo = #SEQ_NUM_WRONG_SIZE
             THEN
               #statStatus := #ERR_SEQ_NUMBER;
               #statSubfunctionStatus := #statRecStruct.backup.SequenceNo;
               #statFBErrorState := #statFBState;
             END_IF;
           ELSIF #instRdRec.ERROR = TRUE THEN
             #statStatus := #ERR_RDREC_VERIFY;
             #statSubfunctionStatus := #instRdRec.STATUS;
             #statFBErrorState := #statFBState;
           END_IF;
         END_REGION verify

       ELSE // Undefined state in state machine reached
         REGION undefined state
           #statStatus := #ERR_UNDEFINED_STATE;
         END_REGION undefined state no relevant case, ready for new request
     END_CASE;
   END_REGION

   REGION OUTPUTS
     // Write outputs
     IF (#statStatus = #STATUS_EXECUTION_FINISHED) AND (#statDone = FALSE) THEN // Execution finished without errors
       REGION execution finished
         #statDone := TRUE;
         #statBusy := FALSE;
         #statError := FALSE;
         #len := #statLen;
         // execution aborted --> set state no processing
         #statFBState := #FB_STATE_NO_PROCESSING;
       END_REGION execution finished

     ELSIF (#statStatus.%X15 = TRUE) AND (#statError = FALSE) THEN // Error occurred (#statStatus is 16#8000 to 16#FFFF)
       REGION error occured
         #statDone := FALSE;
         #statBusy := FALSE;
         #statError := TRUE;
         // Write diagnostics
         #diagnostics.status := #statStatus;
         #diagnostics.subfunctionStatus := #statSubfunctionStatus;
         #diagnostics.stateNumber := #statFBErrorState;
         // Call instructions with FALSE to be ready for next job
         #instRdRec(REQ    := FALSE,
                    RECORD := #statRecStruct.backup);

         #instWrRec(REQ := FALSE);
         // execution aborted --> set state no processing
         #statFBState := #FB_STATE_NO_PROCESSING;
       END_REGION error occured

     ELSIF (#tempExecute = FALSE) AND ((#statDone = TRUE) OR (#statError = TRUE)) THEN // Reset outputs
       REGION execute reset
         #statDone := FALSE;
         #statBusy := FALSE;
         #statError := FALSE;
         #statStatus := #STATUS_NO_CALL;
         #len := 0;
       END_REGION execute reset
     END_IF;

     REGION write static values to outputs
       #done := #statDone;
       #busy := #statBusy;
       #error := #statError;
       #status := #statStatus;
       ENO := NOT #statError;
     END_REGION write static values to outputs
   END_REGION OUTPUTS
END_FUNCTION_BLOCK

// folder: Device-specific blocks/SIMATIC RF200

